Fanuc KAREL source: kt00068.KL

-- PROVISIONAL review KL for V770-1; original PC SHA256 19381a18d174ad5d02bfbcc66b5af76ac4df5f6d21851a1db454b0962bfef074
-- Incomplete behavior may be omitted. Consult companion uncertainty JSON. Do not deploy.
PROGRAM KT00068
%NOLOCKGROUP
VAR
  I1 : INTEGER
  R2 : REAL
  OUT : REAL
BEGIN
  -- UNRESOLVED_PC offsets 5-16; opcodes 2E,23
  -- UNRESOLVED_PC offsets 21-32; opcodes 2E,23
  -- UNRESOLVED_PC offsets 37-58; opcodes 21,21,29,64,6B,23
  -- UNRESOLVED_PC offsets 63-67; opcodes 7F
END KT00068
